(*
SPDX-FileCopyrightText: c 2026 Oleksandr Tiutyk <trofimich@gmail.com>
SPDX-License-Identifier: MIT
License: https://opensource.org/license/mit
*)

(*!
<summary>Checks raw membership for a present value, a duplicate and an absent value.</summary>
<description>
Borrows a group-owned list reserved for this case. Use from one task at a stable address.
Teardown clears the list before publication.
</description>
*)

{attribute 'no_assign'}
{attribute 'no_explicit_call' := 'do not call this function block directly'}
FUNCTION_BLOCK ListContainsTest EXTENDS TOF_Testing.SingleCycleTest
VAR_STAT
	{attribute 'hide'}
	_ClassName : STRING := __POUNAME();
END_VAR
VAR
	_List : TOF_Collections.IList;
END_VAR

(*!
<summary>Clears the fixture before the runner publishes the result.</summary>
<description>
Also runs after an unexpected exception interrupts the case.
</description>
*)
METHOD PROTECTED AfterTest
_List.Clear();
END_METHOD

//! <summary>Borrows the concrete class name. Callers must not modify it.</summary>
{attribute 'monitoring' := 'call'}
PROPERTY ClassName : REFERENCE TO STRING
GET
ClassName REF= _ClassName;
END_GET
END_PROPERTY

(*!
<summary>Checks raw membership for a present value, a duplicate and an absent value.</summary>
*)
METHOD PROTECTED ExecuteTest
VAR
	values : ARRAY [0..5] OF STRING := ['String0', 'String1', 'String2', 'String3', 'String4', 'String5'];
END_VAR
_List.AppendCopy(value := values[0]);
_List.AppendCopy(value := values[1]);
_List.AppendCopy(value := values[2]);
_List.AppendCopy(value := values[3]);
_List.AppendCopy(value := values[2]);
_List.AppendCopy(value := values[3]);

Assert.ThatBool(
	actual := _List.Contains(value := values[1]),
	message := "Contains must find String1"
).IsTrue();

Assert.ThatBool(
	actual := _List.Contains(value := values[3]),
	message := "Contains must find the duplicated String3"
).IsTrue();

Assert.ThatBool(
	actual := _List.Contains(value := values[5]),
	message := "Contains must reject absent String5"
).IsFalse();

Assert.ThatDInt(
	actual := _List.Length,
	message := "Contains must preserve all entries"
).ToBe(expected := DINT#6);
END_METHOD

(*!
<summary>Binds the list fixture for this case.</summary>
<description>
Stores a borrowed interface without invoking the fixture. The owning group keeps it alive and
reserves it for this case. TestElement initializes the name and parent.
</description>
<param name="name">Display name of this case.</param>
<param name="parent">Group that owns this case.</param>
<param name="list">Required live list reserved for this case.</param>
*)
METHOD FB_init : BOOL
VAR_INPUT
	bInitRetains: BOOL; // TRUE: the retain variables are initialized (reset warm / reset cold)
	bInCopyCode: BOOL; // TRUE: the instance will be copied to the copy code afterward (online change)
	name : WSTRING;
	parent : TOF_Testing.ITestElement;
	list : TOF_Collections.IList;
END_VAR
_List := list;
FB_init := TRUE;
END_METHOD

//! <summary>Borrows the compiler-initialized namespace name. Callers must not modify it.</summary>
{attribute 'monitoring' := 'call'}
PROPERTY NamespaceName : REFERENCE TO STRING
GET
NamespaceName REF= CurrentNamespace.Name;
END_GET
END_PROPERTY

//! <summary>Reports the concrete instance size in bytes.</summary>
{attribute 'monitoring' := 'call'}
PROPERTY SelfSize : ULINT
GET
SelfSize := XSIZEOF(THIS^);
END_GET
END_PROPERTY

END_FUNCTION_BLOCK

(* stored: Version 1.1.0.1, ProductVersion 3.1.4026.21
   POU ListContainsTest: Id {4e572c2b-d3f2-4069-8645-cb9b98b97e19}, SpecialFunc None
   Method AfterTest: Id {22a9a27f-5d98-411a-bf5c-7799bc06cb48}
   Property ClassName: Id {bcc02f0c-9259-440a-ac30-ef24d4aaebcf}
   Get Get: Id {6fa25821-cd78-4169-abca-20e26186231c}
   Method ExecuteTest: Id {0d229432-fe9d-4562-a4bd-df8ea223f500}
   Method FB_init: Id {8cee251b-f924-41e4-8ccd-c87186da2a88}
   Property NamespaceName: Id {e4e4ee70-7fb3-43c3-bbe7-05962ae7d1b8}
   Get Get: Id {94163645-03c3-4151-8911-813a5f6a2fef}
   Property SelfSize: Id {9c1674a6-87c2-45c8-b3b9-37aa9322c16d}
   Get Get: Id {6e286d69-c010-4365-a521-657efb6f199b} *)
